Fanuc KAREL source: KC00062.KL

PROGRAM KC00062
%NOLOCKGROUP
%ENVIRONMENT CVIS
VAR
  I: INTEGER
  J: INTEGER
  K: INTEGER
  R: REAL
  B: BOOLEAN
  S: STRING[80]
  T: STRING[80]
  P: PATH
  Q: PATH
  AI: ARRAY[8] OF INTEGER
  AB: ARRAY[244] OF BYTE
  F: POSITION
BEGIN
  INTSCT_VL_PL(P,F,Q,I)
END KC00062
